(* IEC 61131-3 sources: llm-plc-st-eval/data/definitivo/gemini-3.1-pro-preview/A5/zero_shot, 3 files *)

(* ---- ejec_1.st ---- *)
```iecst
TYPE ST_Evento :
STRUCT
    codigo : INT;   (* Código del evento *)
    marca  : TIME;  (* Tiempo acumulado en el momento del evento *)
END_STRUCT
END_TYPE

FUNCTION_BLOCK FB_Registro
VAR_INPUT
    evento      : INT;      (* Código del evento a registrar *)
    nuevoEvento : BOOL;     (* Disparador para registrar el evento (flanco de subida) *)
    ciclo       : TIME;     (* Período de ejecución del bloque *)
END_VAR

VAR_OUTPUT
    buffer      : ARRAY[0..19] OF ST_Evento; (* Buffer circular de eventos *)
    indice      : INT := -1;                 (* Índice del último evento registrado (-1 si está vacío) *)
    nEventos    : INT := 0;                  (* Cantidad de eventos válidos en el buffer (0 a 20) *)
END_VAR

VAR
    tiempoAcumulado : TIME := T#0s;          (* Tiempo total acumulado desde el arranque *)
    prevNuevoEvento : BOOL := FALSE;         (* Memoria para detectar el flanco de subida *)
END_VAR

(* 1. Acumular el tiempo de ejecución en cada ciclo *)
tiempoAcumulado := tiempoAcumulado + ciclo;

(* 2. Detectar transición de FALSE a TRUE en nuevoEvento *)
IF nuevoEvento AND NOT prevNuevoEvento THEN

    (* 3. Calcular el nuevo índice (buffer circular de 0 a 19) *)
    indice := indice + 1;
    IF indice > 19 THEN
        indice := 0;
    END_IF;

    (* 4. Registrar los datos en el buffer *)
    buffer[indice].codigo := evento;
    buffer[indice].marca  := tiempoAcumulado;

    (* 5. Actualizar la cantidad de eventos válidos (tope en 20) *)
    IF nEventos < 20 THEN
        nEventos := nEventos + 1;
    END_IF;

END_IF;

(* 6. Actualizar la memoria del flanco para el siguiente ciclo *)
prevNuevoEvento := nuevoEvento;

END_FUNCTION_BLOCK
```

(* ---- ejec_2.st ---- *)
```iecst
TYPE ST_Evento :
STRUCT
    codigo : INT;  // Código del evento
    marca  : TIME; // Tiempo acumulado en el momento del evento
END_STRUCT
END_TYPE

FUNCTION_BLOCK FB_Registro
VAR_INPUT
    evento      : INT;  // Código del evento a registrar
    nuevoEvento : BOOL; // Señal para registrar evento (flanco de subida)
    ciclo       : TIME; // Período de ejecución para el tiempo acumulado
END_VAR

VAR_OUTPUT
    buffer      : ARRAY[0..19] OF ST_Evento; // Buffer circular de eventos
    indice      : INT := -1;                 // Posición del último evento (-1 si está vacío)
    nEventos    : INT := 0;                  // Cantidad de eventos válidos (0 a 20)
END_VAR

VAR
    tiempoAcumulado : TIME := T#0s;          // Tiempo total acumulado desde el arranque
    prevNuevoEvento : BOOL := FALSE;         // Memoria para detección de flanco de subida
END_VAR

// 1. Acumular el tiempo de ejecución en cada ciclo
tiempoAcumulado := tiempoAcumulado + ciclo;

// 2. Detectar transición de FALSE a TRUE en nuevoEvento (flanco de subida)
IF nuevoEvento AND NOT prevNuevoEvento THEN

    // 3. Actualizar el índice de forma circular (0 a 19)
    indice := indice + 1;
    IF indice > 19 THEN
        indice := 0;
    END_IF;

    // 4. Registrar el evento en la posición actual del buffer
    buffer[indice].codigo := evento;
    buffer[indice].marca  := tiempoAcumulado;

    // 5. Actualizar el contador de eventos válidos (saturado en 20)
    IF nEventos < 20 THEN
        nEventos := nEventos + 1;
    END_IF;

END_IF;

// 6. Actualizar la memoria del estado anterior para el detector de flanco
prevNuevoEvento := nuevoEvento;

END_FUNCTION_BLOCK
```

(* ---- ejec_3.st ---- *)
```iecst
TYPE ST_Evento :
STRUCT
    codigo : INT;  (* Código del evento *)
    marca  : TIME; (* Tiempo acumulado en el momento del evento *)
END_STRUCT
END_TYPE

FUNCTION_BLOCK FB_Registro
VAR_INPUT
    evento      : INT;  (* Valor del evento a registrar *)
    nuevoEvento : BOOL; (* Señal para registrar un nuevo evento (flanco de subida) *)
    ciclo       : TIME; (* Período de ejecución del bloque *)
END_VAR

VAR_OUTPUT
    buffer      : ARRAY[0..19] OF ST_Evento; (* Arreglo circular de eventos *)
    indice      : INT := -1;                 (* Posición del último evento registrado (-1 si no hay) *)
    nEventos    : INT := 0;                  (* Número de eventos válidos en el buffer (0 a 20) *)
END_VAR

VAR
    tiempoAcumulado : TIME := T#0s;  (* Tiempo acumulado desde el arranque *)
    prevNuevoEvento : BOOL := FALSE; (* Memoria para detectar el flanco de subida *)
END_VAR

(* Acumular el tiempo de ciclo en cada ejecución *)
tiempoAcumulado := tiempoAcumulado + ciclo;

(* Detectar transición de FALSE a TRUE en nuevoEvento *)
IF nuevoEvento AND NOT prevNuevoEvento THEN

    (* Incrementar índice y aplicar lógica de buffer circular *)
    indice := indice + 1;
    IF indice > 19 THEN
        indice := 0;
    END_IF;

    (* Registrar el evento y la marca de tiempo en la posición actual *)
    buffer[indice].codigo := evento;
    buffer[indice].marca  := tiempoAcumulado;

    (* Incrementar el contador de eventos válidos hasta un máximo de 20 *)
    IF nEventos < 20 THEN
        nEventos := nEventos + 1;
    END_IF;

END_IF;

(* Guardar el estado actual para la detección de flanco en el próximo ciclo *)
prevNuevoEvento := nuevoEvento;

END_FUNCTION_BLOCK
```
